(* IEC 61131-3 sources: virtual-bottling-plant/plc/src/generated/alarms, 1 file *)

(* ---- FB_AlarmTable.st ---- *)
(* GENERATED by plc/scripts/gen_plc_io.py from contracts/modbus/plc-io.yaml. Do not edit by hand. *)
(* Line 1 alarm table. *)
FUNCTION_BLOCK FB_AlarmTable
  VAR_INPUT
    AckId : INT; (* alarm id, -1 = all, 0 = none *)
    T101_BrixOutOfSpec : BOOL; (* 1, P3: Batch Brix out of tolerance *)
    T101_CommsLost : BOOL; (* 2, P1: T-101 remote I/O not responding *)
    P201_LowTemp : BOOL; (* 3, P1: Outlet below 83 °C *)
    P201_SteamLow : BOOL; (* 4, P2: Steam pressure low *)
    P201_CommsLost : BOOL; (* 5, P1: P-201 remote I/O not responding *)
    T301_LowLevel : BOOL; (* 6, P3: Buffer below filler start level *)
    T301_CommsLost : BOOL; (* 7, P1: T-301 remote I/O not responding *)
    F401_NozzleLeak : BOOL; (* 8, P2: Filler nozzle leak *)
    F401_CommsLost : BOOL; (* 9, P1: F-401 remote I/O not responding *)
    C501_Jam : BOOL; (* 10, P2: Capper jam *)
    C501_Breakdown : BOOL; (* 11, P1: Capper breakdown *)
    C501_CapsEmpty : BOOL; (* 12, P3: Cap hopper empty *)
    C501_CommsLost : BOOL; (* 13, P1: C-501 remote I/O not responding *)
    L601_RollEmpty : BOOL; (* 14, P3: Label roll empty *)
    L601_LabelError : BOOL; (* 15, P2: Label glue / application error *)
    L601_Breakdown : BOOL; (* 16, P1: Labeler breakdown *)
    L601_CommsLost : BOOL; (* 17, P1: L-601 remote I/O not responding *)
    Q701_CommsLost : BOOL; (* 18, P1: Q-701 remote I/O not responding *)
    K801_Jam : BOOL; (* 19, P2: Case packer jam *)
    K801_Breakdown : BOOL; (* 20, P1: Case packer breakdown *)
    K801_CommsLost : BOOL; (* 21, P1: K-801 remote I/O not responding *)
    LINE_CommsLost : BOOL; (* 22, P1: Line I/O (clock *)
  END_VAR
  VAR_OUTPUT
    Summary : ST_AlarmSummary;
  END_VAR
  VAR
    Alm_T101_BrixOutOfSpec : FB_Alarm;
    Alm_T101_CommsLost : FB_Alarm;
    Alm_P201_LowTemp : FB_Alarm;
    Alm_P201_SteamLow : FB_Alarm;
    Alm_P201_CommsLost : FB_Alarm;
    Alm_T301_LowLevel : FB_Alarm;
    Alm_T301_CommsLost : FB_Alarm;
    Alm_F401_NozzleLeak : FB_Alarm;
    Alm_F401_CommsLost : FB_Alarm;
    Alm_C501_Jam : FB_Alarm;
    Alm_C501_Breakdown : FB_Alarm;
    Alm_C501_CapsEmpty : FB_Alarm;
    Alm_C501_CommsLost : FB_Alarm;
    Alm_L601_RollEmpty : FB_Alarm;
    Alm_L601_LabelError : FB_Alarm;
    Alm_L601_Breakdown : FB_Alarm;
    Alm_L601_CommsLost : FB_Alarm;
    Alm_Q701_CommsLost : FB_Alarm;
    Alm_K801_Jam : FB_Alarm;
    Alm_K801_Breakdown : FB_Alarm;
    Alm_K801_CommsLost : FB_Alarm;
    Alm_LINE_CommsLost : FB_Alarm;
    FirstOutFree : BOOL := TRUE;
    Standing : INT;
    StandingLastScan : INT;
  END_VAR
  (* First-out re-arms once every alarm is cleared and acknowledged. The line's
     FirstOutId follows the alarm holding the flag, so it drops to 0 as soon as that
     alarm is cleared and acked, even while other alarms are still shown. *)
  IF StandingLastScan = 0 THEN
    FirstOutFree := TRUE;
  END_IF;
  Summary.FirstOutId := 0;
  Standing := 0;
  Summary.ActiveCount := 0;
  Summary.T101_Word := 0;
  Summary.T101_ActiveId := 0;
  Summary.P201_Word := 0;
  Summary.P201_ActiveId := 0;
  Summary.T301_Word := 0;
  Summary.T301_ActiveId := 0;
  Summary.F401_Word := 0;
  Summary.F401_ActiveId := 0;
  Summary.C501_Word := 0;
  Summary.C501_ActiveId := 0;
  Summary.L601_Word := 0;
  Summary.L601_ActiveId := 0;
  Summary.Q701_Word := 0;
  Summary.Q701_ActiveId := 0;
  Summary.K801_Word := 0;
  Summary.K801_ActiveId := 0;
  Summary.LINE_Word := 0;
  Summary.LINE_ActiveId := 0;
  Alm_T101_BrixOutOfSpec(Condition := T101_BrixOutOfSpec, AckId := AckId, Id := 1, Priority := 3, FirstOutFree := FirstOutFree);
  Summary.W1 := Alm_T101_BrixOutOfSpec.StatusWord;
  IF Alm_T101_BrixOutOfSpec.Active THEN Summary.T101_Word := Summary.T101_Word + 1; Summary.ActiveCount := Summary.ActiveCount + 1; END_IF;
  IF Alm_T101_BrixOutOfSpec.Active AND Summary.T101_ActiveId = 0 THEN Summary.T101_ActiveId := 1; END_IF;
  IF Alm_T101_BrixOutOfSpec.Shown THEN Standing := Standing + 1; END_IF;
  IF Alm_T101_BrixOutOfSpec.FirstOut THEN Summary.FirstOutId := 1; END_IF;
  Alm_T101_CommsLost(Condition := T101_CommsLost, AckId := AckId, Id := 2, Priority := 1, FirstOutFree := FirstOutFree);
  Summary.W2 := Alm_T101_CommsLost.StatusWord;
  IF Alm_T101_CommsLost.Active THEN Summary.T101_Word := Summary.T101_Word + 2; Summary.ActiveCount := Summary.ActiveCount + 1; END_IF;
  IF Alm_T101_CommsLost.Active AND Summary.T101_ActiveId = 0 THEN Summary.T101_ActiveId := 2; END_IF;
  IF Alm_T101_CommsLost.Shown THEN Standing := Standing + 1; END_IF;
  IF Alm_T101_CommsLost.FirstOut THEN Summary.FirstOutId := 2; END_IF;
  Alm_P201_LowTemp(Condition := P201_LowTemp, AckId := AckId, Id := 3, Priority := 1, FirstOutFree := FirstOutFree);
  Summary.W3 := Alm_P201_LowTemp.StatusWord;
  IF Alm_P201_LowTemp.Active THEN Summary.P201_Word := Summary.P201_Word + 1; Summary.ActiveCount := Summary.ActiveCount + 1; END_IF;
  IF Alm_P201_LowTemp.Active AND Summary.P201_ActiveId = 0 THEN Summary.P201_ActiveId := 3; END_IF;
  IF Alm_P201_LowTemp.Shown THEN Standing := Standing + 1; END_IF;
  IF Alm_P201_LowTemp.FirstOut THEN Summary.FirstOutId := 3; END_IF;
  Alm_P201_SteamLow(Condition := P201_SteamLow, AckId := AckId, Id := 4, Priority := 2, FirstOutFree := FirstOutFree);
  Summary.W4 := Alm_P201_SteamLow.StatusWord;
  IF Alm_P201_SteamLow.Active THEN Summary.P201_Word := Summary.P201_Word + 2; Summary.ActiveCount := Summary.ActiveCount + 1; END_IF;
  IF Alm_P201_SteamLow.Active AND Summary.P201_ActiveId = 0 THEN Summary.P201_ActiveId := 4; END_IF;
  IF Alm_P201_SteamLow.Shown THEN Standing := Standing + 1; END_IF;
  IF Alm_P201_SteamLow.FirstOut THEN Summary.FirstOutId := 4; END_IF;
  Alm_P201_CommsLost(Condition := P201_CommsLost, AckId := AckId, Id := 5, Priority := 1, FirstOutFree := FirstOutFree);
  Summary.W5 := Alm_P201_CommsLost.StatusWord;
  IF Alm_P201_CommsLost.Active THEN Summary.P201_Word := Summary.P201_Word + 4; Summary.ActiveCount := Summary.ActiveCount + 1; END_IF;
  IF Alm_P201_CommsLost.Active AND Summary.P201_ActiveId = 0 THEN Summary.P201_ActiveId := 5; END_IF;
  IF Alm_P201_CommsLost.Shown THEN Standing := Standing + 1; END_IF;
  IF Alm_P201_CommsLost.FirstOut THEN Summary.FirstOutId := 5; END_IF;
  Alm_T301_LowLevel(Condition := T301_LowLevel, AckId := AckId, Id := 6, Priority := 3, FirstOutFree := FirstOutFree);
  Summary.W6 := Alm_T301_LowLevel.StatusWord;
  IF Alm_T301_LowLevel.Active THEN Summary.T301_Word := Summary.T301_Word + 1; Summary.ActiveCount := Summary.ActiveCount + 1; END_IF;
  IF Alm_T301_LowLevel.Active AND Summary.T301_ActiveId = 0 THEN Summary.T301_ActiveId := 6; END_IF;
  IF Alm_T301_LowLevel.Shown THEN Standing := Standing + 1; END_IF;
  IF Alm_T301_LowLevel.FirstOut THEN Summary.FirstOutId := 6; END_IF;
  Alm_T301_CommsLost(Condition := T301_CommsLost, AckId := AckId, Id := 7, Priority := 1, FirstOutFree := FirstOutFree);
  Summary.W7 := Alm_T301_CommsLost.StatusWord;
  IF Alm_T301_CommsLost.Active THEN Summary.T301_Word := Summary.T301_Word + 2; Summary.ActiveCount := Summary.ActiveCount + 1; END_IF;
  IF Alm_T301_CommsLost.Active AND Summary.T301_ActiveId = 0 THEN Summary.T301_ActiveId := 7; END_IF;
  IF Alm_T301_CommsLost.Shown THEN Standing := Standing + 1; END_IF;
  IF Alm_T301_CommsLost.FirstOut THEN Summary.FirstOutId := 7; END_IF;
  Alm_F401_NozzleLeak(Condition := F401_NozzleLeak, AckId := AckId, Id := 8, Priority := 2, FirstOutFree := FirstOutFree);
  Summary.W8 := Alm_F401_NozzleLeak.StatusWord;
  IF Alm_F401_NozzleLeak.Active THEN Summary.F401_Word := Summary.F401_Word + 1; Summary.ActiveCount := Summary.ActiveCount + 1; END_IF;
  IF Alm_F401_NozzleLeak.Active AND Summary.F401_ActiveId = 0 THEN Summary.F401_ActiveId := 8; END_IF;
  IF Alm_F401_NozzleLeak.Shown THEN Standing := Standing + 1; END_IF;
  IF Alm_F401_NozzleLeak.FirstOut THEN Summary.FirstOutId := 8; END_IF;
  Alm_F401_CommsLost(Condition := F401_CommsLost, AckId := AckId, Id := 9, Priority := 1, FirstOutFree := FirstOutFree);
  Summary.W9 := Alm_F401_CommsLost.StatusWord;
  IF Alm_F401_CommsLost.Active THEN Summary.F401_Word := Summary.F401_Word + 2; Summary.ActiveCount := Summary.ActiveCount + 1; END_IF;
  IF Alm_F401_CommsLost.Active AND Summary.F401_ActiveId = 0 THEN Summary.F401_ActiveId := 9; END_IF;
  IF Alm_F401_CommsLost.Shown THEN Standing := Standing + 1; END_IF;
  IF Alm_F401_CommsLost.FirstOut THEN Summary.FirstOutId := 9; END_IF;
  Alm_C501_Jam(Condition := C501_Jam, AckId := AckId, Id := 10, Priority := 2, FirstOutFree := FirstOutFree);
  Summary.W10 := Alm_C501_Jam.StatusWord;
  IF Alm_C501_Jam.Active THEN Summary.C501_Word := Summary.C501_Word + 1; Summary.ActiveCount := Summary.ActiveCount + 1; END_IF;
  IF Alm_C501_Jam.Active AND Summary.C501_ActiveId = 0 THEN Summary.C501_ActiveId := 10; END_IF;
  IF Alm_C501_Jam.Shown THEN Standing := Standing + 1; END_IF;
  IF Alm_C501_Jam.FirstOut THEN Summary.FirstOutId := 10; END_IF;
  Alm_C501_Breakdown(Condition := C501_Breakdown, AckId := AckId, Id := 11, Priority := 1, FirstOutFree := FirstOutFree);
  Summary.W11 := Alm_C501_Breakdown.StatusWord;
  IF Alm_C501_Breakdown.Active THEN Summary.C501_Word := Summary.C501_Word + 2; Summary.ActiveCount := Summary.ActiveCount + 1; END_IF;
  IF Alm_C501_Breakdown.Active AND Summary.C501_ActiveId = 0 THEN Summary.C501_ActiveId := 11; END_IF;
  IF Alm_C501_Breakdown.Shown THEN Standing := Standing + 1; END_IF;
  IF Alm_C501_Breakdown.FirstOut THEN Summary.FirstOutId := 11; END_IF;
  Alm_C501_CapsEmpty(Condition := C501_CapsEmpty, AckId := AckId, Id := 12, Priority := 3, FirstOutFree := FirstOutFree);
  Summary.W12 := Alm_C501_CapsEmpty.StatusWord;
  IF Alm_C501_CapsEmpty.Active THEN Summary.C501_Word := Summary.C501_Word + 4; Summary.ActiveCount := Summary.ActiveCount + 1; END_IF;
  IF Alm_C501_CapsEmpty.Active AND Summary.C501_ActiveId = 0 THEN Summary.C501_ActiveId := 12; END_IF;
  IF Alm_C501_CapsEmpty.Shown THEN Standing := Standing + 1; END_IF;
  IF Alm_C501_CapsEmpty.FirstOut THEN Summary.FirstOutId := 12; END_IF;
  Alm_C501_CommsLost(Condition := C501_CommsLost, AckId := AckId, Id := 13, Priority := 1, FirstOutFree := FirstOutFree);
  Summary.W13 := Alm_C501_CommsLost.StatusWord;
  IF Alm_C501_CommsLost.Active THEN Summary.C501_Word := Summary.C501_Word + 8; Summary.ActiveCount := Summary.ActiveCount + 1; END_IF;
  IF Alm_C501_CommsLost.Active AND Summary.C501_ActiveId = 0 THEN Summary.C501_ActiveId := 13; END_IF;
  IF Alm_C501_CommsLost.Shown THEN Standing := Standing + 1; END_IF;
  IF Alm_C501_CommsLost.FirstOut THEN Summary.FirstOutId := 13; END_IF;
  Alm_L601_RollEmpty(Condition := L601_RollEmpty, AckId := AckId, Id := 14, Priority := 3, FirstOutFree := FirstOutFree);
  Summary.W14 := Alm_L601_RollEmpty.StatusWord;
  IF Alm_L601_RollEmpty.Active THEN Summary.L601_Word := Summary.L601_Word + 1; Summary.ActiveCount := Summary.ActiveCount + 1; END_IF;
  IF Alm_L601_RollEmpty.Active AND Summary.L601_ActiveId = 0 THEN Summary.L601_ActiveId := 14; END_IF;
  IF Alm_L601_RollEmpty.Shown THEN Standing := Standing + 1; END_IF;
  IF Alm_L601_RollEmpty.FirstOut THEN Summary.FirstOutId := 14; END_IF;
  Alm_L601_LabelError(Condition := L601_LabelError, AckId := AckId, Id := 15, Priority := 2, FirstOutFree := FirstOutFree);
  Summary.W15 := Alm_L601_LabelError.StatusWord;
  IF Alm_L601_LabelError.Active THEN Summary.L601_Word := Summary.L601_Word + 2; Summary.ActiveCount := Summary.ActiveCount + 1; END_IF;
  IF Alm_L601_LabelError.Active AND Summary.L601_ActiveId = 0 THEN Summary.L601_ActiveId := 15; END_IF;
  IF Alm_L601_LabelError.Shown THEN Standing := Standing + 1; END_IF;
  IF Alm_L601_LabelError.FirstOut THEN Summary.FirstOutId := 15; END_IF;
  Alm_L601_Breakdown(Condition := L601_Breakdown, AckId := AckId, Id := 16, Priority := 1, FirstOutFree := FirstOutFree);
  Summary.W16 := Alm_L601_Breakdown.StatusWord;
  IF Alm_L601_Breakdown.Active THEN Summary.L601_Word := Summary.L601_Word + 4; Summary.ActiveCount := Summary.ActiveCount + 1; END_IF;
  IF Alm_L601_Breakdown.Active AND Summary.L601_ActiveId = 0 THEN Summary.L601_ActiveId := 16; END_IF;
  IF Alm_L601_Breakdown.Shown THEN Standing := Standing + 1; END_IF;
  IF Alm_L601_Breakdown.FirstOut THEN Summary.FirstOutId := 16; END_IF;
  Alm_L601_CommsLost(Condition := L601_CommsLost, AckId := AckId, Id := 17, Priority := 1, FirstOutFree := FirstOutFree);
  Summary.W17 := Alm_L601_CommsLost.StatusWord;
  IF Alm_L601_CommsLost.Active THEN Summary.L601_Word := Summary.L601_Word + 8; Summary.ActiveCount := Summary.ActiveCount + 1; END_IF;
  IF Alm_L601_CommsLost.Active AND Summary.L601_ActiveId = 0 THEN Summary.L601_ActiveId := 17; END_IF;
  IF Alm_L601_CommsLost.Shown THEN Standing := Standing + 1; END_IF;
  IF Alm_L601_CommsLost.FirstOut THEN Summary.FirstOutId := 17; END_IF;
  Alm_Q701_CommsLost(Condition := Q701_CommsLost, AckId := AckId, Id := 18, Priority := 1, FirstOutFree := FirstOutFree);
  Summary.W18 := Alm_Q701_CommsLost.StatusWord;
  IF Alm_Q701_CommsLost.Active THEN Summary.Q701_Word := Summary.Q701_Word + 1; Summary.ActiveCount := Summary.ActiveCount + 1; END_IF;
  IF Alm_Q701_CommsLost.Active AND Summary.Q701_ActiveId = 0 THEN Summary.Q701_ActiveId := 18; END_IF;
  IF Alm_Q701_CommsLost.Shown THEN Standing := Standing + 1; END_IF;
  IF Alm_Q701_CommsLost.FirstOut THEN Summary.FirstOutId := 18; END_IF;
  Alm_K801_Jam(Condition := K801_Jam, AckId := AckId, Id := 19, Priority := 2, FirstOutFree := FirstOutFree);
  Summary.W19 := Alm_K801_Jam.StatusWord;
  IF Alm_K801_Jam.Active THEN Summary.K801_Word := Summary.K801_Word + 1; Summary.ActiveCount := Summary.ActiveCount + 1; END_IF;
  IF Alm_K801_Jam.Active AND Summary.K801_ActiveId = 0 THEN Summary.K801_ActiveId := 19; END_IF;
  IF Alm_K801_Jam.Shown THEN Standing := Standing + 1; END_IF;
  IF Alm_K801_Jam.FirstOut THEN Summary.FirstOutId := 19; END_IF;
  Alm_K801_Breakdown(Condition := K801_Breakdown, AckId := AckId, Id := 20, Priority := 1, FirstOutFree := FirstOutFree);
  Summary.W20 := Alm_K801_Breakdown.StatusWord;
  IF Alm_K801_Breakdown.Active THEN Summary.K801_Word := Summary.K801_Word + 2; Summary.ActiveCount := Summary.ActiveCount + 1; END_IF;
  IF Alm_K801_Breakdown.Active AND Summary.K801_ActiveId = 0 THEN Summary.K801_ActiveId := 20; END_IF;
  IF Alm_K801_Breakdown.Shown THEN Standing := Standing + 1; END_IF;
  IF Alm_K801_Breakdown.FirstOut THEN Summary.FirstOutId := 20; END_IF;
  Alm_K801_CommsLost(Condition := K801_CommsLost, AckId := AckId, Id := 21, Priority := 1, FirstOutFree := FirstOutFree);
  Summary.W21 := Alm_K801_CommsLost.StatusWord;
  IF Alm_K801_CommsLost.Active THEN Summary.K801_Word := Summary.K801_Word + 4; Summary.ActiveCount := Summary.ActiveCount + 1; END_IF;
  IF Alm_K801_CommsLost.Active AND Summary.K801_ActiveId = 0 THEN Summary.K801_ActiveId := 21; END_IF;
  IF Alm_K801_CommsLost.Shown THEN Standing := Standing + 1; END_IF;
  IF Alm_K801_CommsLost.FirstOut THEN Summary.FirstOutId := 21; END_IF;
  Alm_LINE_CommsLost(Condition := LINE_CommsLost, AckId := AckId, Id := 22, Priority := 1, FirstOutFree := FirstOutFree);
  Summary.W22 := Alm_LINE_CommsLost.StatusWord;
  IF Alm_LINE_CommsLost.Active THEN Summary.LINE_Word := Summary.LINE_Word + 1; Summary.ActiveCount := Summary.ActiveCount + 1; END_IF;
  IF Alm_LINE_CommsLost.Active AND Summary.LINE_ActiveId = 0 THEN Summary.LINE_ActiveId := 22; END_IF;
  IF Alm_LINE_CommsLost.Shown THEN Standing := Standing + 1; END_IF;
  IF Alm_LINE_CommsLost.FirstOut THEN Summary.FirstOutId := 22; END_IF;

  StandingLastScan := Standing;
END_FUNCTION_BLOCK
